// TIA Portal V19 export
TYPE "EM02_Output"
   STRUCT
      Status : "EM_Output";
      VacuumActive : Bool;
      VacuumBroken : Bool;
   END_STRUCT;
END_TYPE
